(* IEC 61131-3 sources: kkh_knowHow_dgtt/tools/fmse/plc_lib (part 2) *)

(* ---- FB_SafetyCoupling.st ---- *)
(*==================================================================================================================
  FB_SafetyCoupling  -  safety coupling to the neighbour module (e-stop in + zone free)
  ----------------------------------------------------------------------------------------------------------------
  Library   : FMSE device FB library (item 10A)              Version : 1.0.0 (2026-11-15)
  Rule      : tools/fmse/examples/item10a_examples.json  _rules.fb_library (= 2 x FB_Safe2Ch)
  Codegen   : item 8 pattern COUPLING -> st_codegen.py calls this FB (x<Signal> / q<Signal>)
  Purpose   : Item 8 COUPLING: one FB_Safe2Ch for the e-stop chain coming in, one for the zone-free signal of
              the neighbour. The outputs EstopOut / EnableOut are F-outputs written only by the F-program.
  Interface :
    dir  name                type          default   meaning
    IN   xEstopIn            BOOL          -         e-stop in channel 1 F-copy
    IN   xEstopIn2           BOOL          -         e-stop in channel 2 F-copy
    IN   xZoneFree           BOOL          -         zone free channel 1 F-copy
    IN   xZoneFree2          BOOL          -         zone free channel 2 F-copy
    IN   xReset              BOOL          -         fault reset, rising edge
    CFG  tDisc_ms            DINT          500       discrepancy time [ms]
    OUT  xEstopOk            BOOL          -         e-stop chain closed and reset
    OUT  xZoneOk             BOOL          -         neighbour zone free and reset
    OUT  xResetReq           BOOL          -         one of the two waits for a reset
    OUT  xDiscErr            BOOL          -         discrepancy in one of the two
    OUT  iAlarm              INT           -         local alarm code (0 = none)
  Alarms    : iAlarm = local code a ; Admin.AlarmNo = M*1000 + 10*i + a (decision D2), class per module (D3)
    1  e-stop coupling discrepancy
    2  zone-free coupling discrepancy
  Timing    : Times are counted in calls: n * GC_CYCLE_MS >= t_ms (GC_CYCLE_MS = 100 ms = test bench, TYPES.st).
              In the 10 ms main task set GC_CYCLE_MS := 10 (same behaviour, 10 ms resolution) or replace a counter
              by a TON: ton(IN := <condition>, PT := T#2s); IF ton.Q THEN ... (one call later than the counter).
  Siemens   : SCL (TIA Portal): the same statements; local names are written with '#' (#xRst), the VAR section is
              VAR (STAT) of an FB with an instance DB, R_TRIG / TON are multi-instances, enumerations become INT
              constants (E_DriveState.FAULT -> 9), MIN / LIMIT exist, '16#0080' is written W#16#80 for a WORD.
  NOTICE    : ALL VALUES ARE EXAMPLES. Real PLC code is written, reviewed, tested and signed off by qualified
              people. Safety functions only in the F-program; this FB only reads F-copies and writes no F-signal.
==================================================================================================================*)
FUNCTION_BLOCK FB_SafetyCoupling
VAR_INPUT  (* signals *)
  xEstopIn : BOOL;                          (* e-stop in channel 1 F-copy *)
  xEstopIn2 : BOOL;                         (* e-stop in channel 2 F-copy *)
  xZoneFree : BOOL;                         (* zone free channel 1 F-copy *)
  xZoneFree2 : BOOL;                        (* zone free channel 2 F-copy *)
  xReset : BOOL;                            (* fault reset, rising edge *)
END_VAR
VAR_INPUT  (* configuration (set once, defaults = example values) *)
  tDisc_ms : DINT := 500;                   (* discrepancy time [ms] *)
END_VAR
VAR_OUTPUT  (* outputs *)
  xEstopOk : BOOL;                          (* e-stop chain closed and reset *)
  xZoneOk : BOOL;                           (* neighbour zone free and reset *)
  xResetReq : BOOL;                         (* one of the two waits for a reset *)
  xDiscErr : BOOL;                          (* discrepancy in one of the two *)
  iAlarm : INT;                             (* local alarm code (0 = none) *)
END_VAR
VAR  (* internal *)
  fbEstop : FB_Safe2Ch;                     (* e-stop in *)
  fbZone : FB_Safe2Ch;                      (* zone free *)
END_VAR
fbEstop(xCh1 := xEstopIn, xCh2 := xEstopIn2, xReset := xReset, tDisc_ms := tDisc_ms);
fbZone(xCh1 := xZoneFree, xCh2 := xZoneFree2, xReset := xReset, tDisc_ms := tDisc_ms);
xEstopOk := fbEstop.xOk;
xZoneOk := fbZone.xOk;
xResetReq := fbEstop.xResetReq OR fbZone.xResetReq;
xDiscErr := fbEstop.xDiscErr OR fbZone.xDiscErr;
IF fbEstop.xDiscErr THEN
  iAlarm := 1;                                (* e-stop coupling discrepancy *)
ELSIF fbZone.xDiscErr THEN
  iAlarm := 2;                                (* zone-free coupling discrepancy *)
ELSE
  iAlarm := 0;
END_IF
END_FUNCTION_BLOCK

(* ---- FB_SafeValve.st ---- *)
(*==================================================================================================================
  FB_SafeValve  -  redundant safety valve pair with position feedback
  ----------------------------------------------------------------------------------------------------------------
  Library   : FMSE device FB library (item 10A)              Version : 1.0.0 (2026-11-15)
  Rule      : tools/fmse/examples/item10a_examples.json  _rules.fb_library (= 2 x FB_Edm, bInverted FALSE)
  Codegen   : item 8 pattern SAFE_VALVE -> st_codegen.py calls this FB (x<Signal> / q<Signal>)
  Purpose   : Item 8 SAFE_VALVE: two valves (F-outputs ValveA / ValveB written only by the F-program), each
              with a position switch TRUE = open; FB_Edm with bInverted FALSE checks that each follows.
  Interface :
    dir  name                type          default   meaning
    IN   xCmdA               BOOL          -         F-copy of the F-output ValveA
    IN   xCmdB               BOOL          -         F-copy of the F-output ValveB
    IN   xFbA                BOOL          -         valve A open (DI)
    IN   xFbB                BOOL          -         valve B open (DI)
    IN   xReset              BOOL          -         fault reset, rising edge
    CFG  tEdm_ms             DINT          300       feedback time [ms]
    OUT  xOnA                BOOL          -         valve A open and feedback ok
    OUT  xOnB                BOOL          -         valve B open and feedback ok
    OUT  xError              BOOL          -         error latched (see alarms)
    OUT  iAlarm              INT           -         local alarm code (0 = none)
  Alarms    : iAlarm = local code a ; Admin.AlarmNo = M*1000 + 10*i + a (decision D2), class per module (D3)
    1  valve A feedback does not follow
    2  valve B feedback does not follow
  Timing    : Times are counted in calls: n * GC_CYCLE_MS >= t_ms (GC_CYCLE_MS = 100 ms = test bench, TYPES.st).
              In the 10 ms main task set GC_CYCLE_MS := 10 (same behaviour, 10 ms resolution) or replace a counter
              by a TON: ton(IN := <condition>, PT := T#2s); IF ton.Q THEN ... (one call later than the counter).
  Siemens   : SCL (TIA Portal): the same statements; local names are written with '#' (#xRst), the VAR section is
              VAR (STAT) of an FB with an instance DB, R_TRIG / TON are multi-instances, enumerations become INT
              constants (E_DriveState.FAULT -> 9), MIN / LIMIT exist, '16#0080' is written W#16#80 for a WORD.
  NOTICE    : ALL VALUES ARE EXAMPLES. Real PLC code is written, reviewed, tested and signed off by qualified
              people. Safety functions only in the F-program; this FB only reads F-copies and writes no F-signal.
==================================================================================================================*)
FUNCTION_BLOCK FB_SafeValve
VAR_INPUT  (* signals *)
  xCmdA : BOOL;                             (* F-copy of the F-output ValveA *)
  xCmdB : BOOL;                             (* F-copy of the F-output ValveB *)
  xFbA : BOOL;                              (* valve A open (DI) *)
  xFbB : BOOL;                              (* valve B open (DI) *)
  xReset : BOOL;                            (* fault reset, rising edge *)
END_VAR
VAR_INPUT  (* configuration (set once, defaults = example values) *)
  tEdm_ms : DINT := 300;                    (* feedback time [ms] *)
END_VAR
VAR_OUTPUT  (* outputs *)
  xOnA : BOOL;                              (* valve A open and feedback ok *)
  xOnB : BOOL;                              (* valve B open and feedback ok *)
  xError : BOOL;                            (* error latched (see alarms) *)
  iAlarm : INT;                             (* local alarm code (0 = none) *)
END_VAR
VAR  (* internal *)
  fbA : FB_Edm;                             (* EDM valve A *)
  fbB : FB_Edm;                             (* EDM valve B *)
END_VAR
fbA(xCmd := xCmdA, xFb := xFbA, xReset := xReset, tEdm_ms := tEdm_ms, bInverted := FALSE);
fbB(xCmd := xCmdB, xFb := xFbB, xReset := xReset, tEdm_ms := tEdm_ms, bInverted := FALSE);
xOnA := fbA.xOn;
xOnB := fbB.xOn;
xError := fbA.xError OR fbB.xError;
IF fbA.xError THEN
  iAlarm := 1;                                (* valve A feedback *)
ELSIF fbB.xError THEN
  iAlarm := 2;                                (* valve B feedback *)
ELSE
  iAlarm := 0;
END_IF
END_FUNCTION_BLOCK

(* ---- FB_Scanner.st ---- *)
(*==================================================================================================================
  FB_Scanner  -  safety laser scanner: field-set switching and OSSD mirror
  ----------------------------------------------------------------------------------------------------------------
  Library   : FMSE device FB library (item 10A)              Version : 1.0.0 (2026-11-15)
  Rule      : tools/fmse/examples/item10a_examples.json  _rules.FB_Scanner
  Codegen   : item 8 pattern SCANNER -> st_codegen.py calls this FB (x<Signal> / q<Signal>)
  Purpose   : The standard program selects the field set (the scanner checks the combination); the OSSD pair
              and the warning field are mirrored for diagnosis and HMI.
  Interface :
    dir  name                type          default   meaning
    IN   xOssd1              BOOL          -         OSSD 1 F-copy (TRUE = free)
    IN   xOssd2              BOOL          -         OSSD 2 F-copy (TRUE = free)
    IN   xWarn               BOOL          -         warning field interrupted (DI)
    IN   iField              INT           1         field set 1 = A, 2 = B
    OUT  qFieldA             BOOL          -         field set A select (DO)
    OUT  qFieldB             BOOL          -         field set B select (DO)
    OUT  xFree               BOOL          -         protective field free
    OUT  xWarnOut            BOOL          -         warning field interrupted
    OUT  iAlarm              INT           -         local alarm code (0 = none)
  Alarms    : iAlarm = local code a ; Admin.AlarmNo = M*1000 + 10*i + a (decision D2), class per module (D3)
    2  invalid field set
  Timing    : Times are counted in calls: n * GC_CYCLE_MS >= t_ms (GC_CYCLE_MS = 100 ms = test bench, TYPES.st).
              In the 10 ms main task set GC_CYCLE_MS := 10 (same behaviour, 10 ms resolution) or replace a counter
              by a TON: ton(IN := <condition>, PT := T#2s); IF ton.Q THEN ... (one call later than the counter).
  Siemens   : SCL (TIA Portal): the same statements; local names are written with '#' (#xRst), the VAR section is
              VAR (STAT) of an FB with an instance DB, R_TRIG / TON are multi-instances, enumerations become INT
              constants (E_DriveState.FAULT -> 9), MIN / LIMIT exist, '16#0080' is written W#16#80 for a WORD.
  NOTICE    : ALL VALUES ARE EXAMPLES. Real PLC code is written, reviewed, tested and signed off by qualified
              people. Safety functions only in the F-program; this FB only reads F-copies and writes no F-signal.
==================================================================================================================*)
FUNCTION_BLOCK FB_Scanner
VAR_INPUT  (* signals *)
  xOssd1 : BOOL;                            (* OSSD 1 F-copy (TRUE = free) *)
  xOssd2 : BOOL;                            (* OSSD 2 F-copy (TRUE = free) *)
  xWarn : BOOL;                             (* warning field interrupted (DI) *)
  iField : INT := 1;                        (* field set 1 = A, 2 = B *)
END_VAR
VAR_OUTPUT  (* outputs *)
  qFieldA : BOOL;                           (* field set A select (DO) *)
  qFieldB : BOOL;                           (* field set B select (DO) *)
  xFree : BOOL;                             (* protective field free *)
  xWarnOut : BOOL;                          (* warning field interrupted *)
  iAlarm : INT;                             (* local alarm code (0 = none) *)
END_VAR
qFieldA := iField = 1;
qFieldB := iField = 2;
xFree := xOssd1 AND xOssd2;
xWarnOut := xWarn;
IF iField = 1 OR iField = 2 THEN
  iAlarm := 0;
ELSE
  iAlarm := 2;                                (* invalid field set *)
END_IF
END_FUNCTION_BLOCK

(* ---- FB_Sensor.st ---- *)
(*==================================================================================================================
  FB_Sensor  -  digital sensor with on / off debounce
  ----------------------------------------------------------------------------------------------------------------
  Library   : FMSE device FB library (item 10A)              Version : 1.0.0 (2026-11-15)
  Rule      : tools/fmse/examples/item10a_examples.json  _rules.FB_Sensor
  Codegen   : item 8 pattern SENSOR -> st_codegen.py calls this FB (x<Signal> / q<Signal>)
  Purpose   : Debounce of a digital sensor: the value follows the input only after it differs for tOn_ms (0 -> 1)
              or tOff_ms (1 -> 0); a shorter bounce is ignored. tOn_ms = tOff_ms = 0: one call delay is not added.
  Interface :
    dir  name                type          default   meaning
    IN   xOn                 BOOL          -         sensor input (DI)
    CFG  tOn_ms              DINT          0         debounce time 0 -> 1 [ms]
    CFG  tOff_ms             DINT          0         debounce time 1 -> 0 [ms]
    OUT  xValue              BOOL          -         debounced value
  Alarms    : iAlarm = local code a ; Admin.AlarmNo = M*1000 + 10*i + a (decision D2), class per module (D3)
    none
  Timing    : Times are counted in calls: n * GC_CYCLE_MS >= t_ms (GC_CYCLE_MS = 100 ms = test bench, TYPES.st).
              In the 10 ms main task set GC_CYCLE_MS := 10 (same behaviour, 10 ms resolution) or replace a counter
              by a TON: ton(IN := <condition>, PT := T#2s); IF ton.Q THEN ... (one call later than the counter).
  Siemens   : SCL (TIA Portal): the same statements; local names are written with '#' (#xRst), the VAR section is
              VAR (STAT) of an FB with an instance DB, R_TRIG / TON are multi-instances, enumerations become INT
              constants (E_DriveState.FAULT -> 9), MIN / LIMIT exist, '16#0080' is written W#16#80 for a WORD.
  NOTICE    : ALL VALUES ARE EXAMPLES. Real PLC code is written, reviewed, tested and signed off by qualified
              people. Safety functions only in the F-program; this FB only reads F-copies and writes no F-signal.
==================================================================================================================*)
FUNCTION_BLOCK FB_Sensor
VAR_INPUT  (* signals *)
  xOn : BOOL;                               (* sensor input (DI) *)
END_VAR
VAR_INPUT  (* configuration (set once, defaults = example values) *)
  tOn_ms : DINT := 0;                       (* debounce time 0 -> 1 [ms] *)
  tOff_ms : DINT := 0;                      (* debounce time 1 -> 0 [ms] *)
END_VAR
VAR_OUTPUT  (* outputs *)
  xValue : BOOL;                            (* debounced value *)
END_VAR
VAR  (* internal *)
  nCnt : DINT;                              (* calls with input <> value *)
  tLim : DINT;                              (* active debounce time *)
END_VAR
IF xOn <> xValue THEN
  nCnt := MIN(nCnt + 1, GC_N_MAX);
  IF xOn THEN
    tLim := tOn_ms;
  ELSE
    tLim := tOff_ms;
  END_IF
  IF nCnt * GC_CYCLE_MS >= tLim THEN
    xValue := xOn;
    nCnt := 0;
  END_IF
ELSE
  nCnt := 0;
END_IF
END_FUNCTION_BLOCK

(* ---- FB_SignalTower.st ---- *)
(*==================================================================================================================
  FB_SignalTower  -  signal tower (stack light) and horn per PackML state and alarm class
  ----------------------------------------------------------------------------------------------------------------
  Library   : FMSE device FB library (item 10A)              Version : 1.0.0 (2026-11-15)
  Rule      : tools/fmse/examples/item10a_examples.json  _rules.FB_SignalTower
  Codegen   : item 8 pattern SIGNAL_TOWER -> st_codegen.py calls this FB (x<Signal> / q<Signal>)
  Purpose   : Colours per IEC 60204-1 10.3 / IEC 60073: red = class A alarm or Aborting/Aborted, yellow = class
              B/C or Stopped/Suspended/Held, green = running states, flashing green = Idle/Complete (ready).
              Horn on a new class A/B alarm until acknowledged or no alarm.
  Interface :
    dir  name                type          default   meaning
    IN   iState              INT           2         PackML state number (2 = Stopped)
    IN   iAlarmClass         INT           -         0 none, 1 A, 2 B, 3 C (FB_AlarmMgr)
    IN   xHornAck            BOOL          -         horn acknowledge, rising edge
    OUT  qRed                BOOL          -         red lamp (DO)
    OUT  qYellow             BOOL          -         yellow lamp (DO)
    OUT  qGreen              BOOL          -         green lamp (DO)
    OUT  qBuzzer             BOOL          -         horn (DO)
  Alarms    : iAlarm = local code a ; Admin.AlarmNo = M*1000 + 10*i + a (decision D2), class per module (D3)
    none
  Timing    : Times are counted in calls: n * GC_CYCLE_MS >= t_ms (GC_CYCLE_MS = 100 ms = test bench, TYPES.st).
              In the 10 ms main task set GC_CYCLE_MS := 10 (same behaviour, 10 ms resolution) or replace a counter
              by a TON: ton(IN := <condition>, PT := T#2s); IF ton.Q THEN ... (one call later than the counter).
  Siemens   : SCL (TIA Portal): the same statements; local names are written with '#' (#xRst), the VAR section is
              VAR (STAT) of an FB with an instance DB, R_TRIG / TON are multi-instances, enumerations become INT
              constants (E_DriveState.FAULT -> 9), MIN / LIMIT exist, '16#0080' is written W#16#80 for a WORD.
  NOTICE    : ALL VALUES ARE EXAMPLES. Real PLC code is written, reviewed, tested and signed off by qualified
              people. Safety functions only in the F-program; this FB only reads F-copies and writes no F-signal.
==================================================================================================================*)
FUNCTION_BLOCK FB_SignalTower
VAR_INPUT  (* signals *)
  iState : INT := 2;                        (* PackML state number (2 = Stopped) *)
  iAlarmClass : INT;                        (* 0 none, 1 A, 2 B, 3 C (FB_AlarmMgr) *)
  xHornAck : BOOL;                          (* horn acknowledge, rising edge *)
END_VAR
VAR_OUTPUT  (* outputs *)
  qRed : BOOL;                              (* red lamp (DO) *)
  qYellow : BOOL;                           (* yellow lamp (DO) *)
  qGreen : BOOL;                            (* green lamp (DO) *)
  qBuzzer : BOOL;                           (* horn (DO) *)
END_VAR
VAR  (* internal *)
  nBlink : DINT;                            (* blink counter 0 .. 2*nHalf-1 *)
  nHalf : DINT;                             (* calls per half period *)
  xBlink : BOOL;                            (* 1 Hz blink, TRUE in the first half *)
  rtAck : R_TRIG;                           (* edge of xHornAck *)
  iPrevClass : INT;                         (* alarm class of the last call *)
  xHorn : BOOL;                             (* horn latch *)
END_VAR
nHalf := GC_BLINK_HALF_MS / GC_CYCLE_MS;     (* 5 calls at 100 ms = 1 Hz *)
xBlink := nBlink < nHalf;
nBlink := (nBlink + 1) MOD (2 * nHalf);
rtAck(CLK := xHornAck);
qRed := (iAlarmClass = E_AlarmClass.A) OR (iState = E_PackMLState.ABORTING) OR (iState = E_PackMLState.ABORTED);
qYellow := (iAlarmClass = E_AlarmClass.B) OR (iAlarmClass = E_AlarmClass.C) OR (iState = E_PackMLState.STOPPED)
           OR (iState = E_PackMLState.SUSPENDED) OR (iState = E_PackMLState.HELD);
CASE iState OF
  E_PackMLState.STARTING, E_PackMLState.EXECUTE, E_PackMLState.UNHOLDING, E_PackMLState.UNSUSPENDING,
  E_PackMLState.COMPLETING:
    qGreen := TRUE;
  E_PackMLState.IDLE, E_PackMLState.COMPLETE:
    qGreen := xBlink;                         (* flashing green = ready, waiting *)
ELSE
  qGreen := FALSE;
END_CASE
IF (iAlarmClass = E_AlarmClass.A OR iAlarmClass = E_AlarmClass.B) AND iAlarmClass <> iPrevClass THEN
  xHorn := TRUE;
END_IF
IF rtAck.Q OR iAlarmClass = E_AlarmClass.NONE THEN
  xHorn := FALSE;
END_IF
iPrevClass := iAlarmClass;
qBuzzer := xHorn;
END_FUNCTION_BLOCK

(* ---- FB_TwoHand.st ---- *)
(*==================================================================================================================
  FB_TwoHand  -  diagnostic mirror of a two-hand control (type IIIC)
  ----------------------------------------------------------------------------------------------------------------
  Library   : FMSE device FB library (item 10A)              Version : 1.0.0 (2026-11-15)
  Rule      : tools/fmse/examples/item10a_examples.json  _rules.FB_TwoHand
  Codegen   : item 8 pattern TWOHAND -> st_codegen.py calls this FB (x<Signal> / q<Signal>)
  Purpose   : Two 2-channel buttons, simultaneity 0.5 s (the F-program does the safety function). Pressing the
              second hand later than tSync_ms blocks until both are released. Strict '>': the 5th call (500 ms)
              is still simultaneous.
  Interface :
    dir  name                type          default   meaning
    IN   xLeft               BOOL          -         left button NO (DI)
    IN   xLeft2              BOOL          -         left button NC (DI)
    IN   xRight              BOOL          -         right button NO (DI)
    IN   xRight2             BOOL          -         right button NC (DI)
    CFG  tSync_ms            DINT          500       simultaneity time [ms]
    OUT  xActuated           BOOL          -         both hands, simultaneous
    OUT  xError              BOOL          -         error latched (see alarms)
    OUT  iAlarm              INT           -         local alarm code (0 = none)
  Alarms    : iAlarm = local code a ; Admin.AlarmNo = M*1000 + 10*i + a (decision D2), class per module (D3)
    1  not simultaneous - release both
  Timing    : Times are counted in calls: n * GC_CYCLE_MS >= t_ms (GC_CYCLE_MS = 100 ms = test bench, TYPES.st).
              In the 10 ms main task set GC_CYCLE_MS := 10 (same behaviour, 10 ms resolution) or replace a counter
              by a TON: ton(IN := <condition>, PT := T#2s); IF ton.Q THEN ... (one call later than the counter).
  Siemens   : SCL (TIA Portal): the same statements; local names are written with '#' (#xRst), the VAR section is
              VAR (STAT) of an FB with an instance DB, R_TRIG / TON are multi-instances, enumerations become INT
              constants (E_DriveState.FAULT -> 9), MIN / LIMIT exist, '16#0080' is written W#16#80 for a WORD.
  NOTICE    : ALL VALUES ARE EXAMPLES. Real PLC code is written, reviewed, tested and signed off by qualified
              people. Safety functions only in the F-program; this FB only reads F-copies and writes no F-signal.
==================================================================================================================*)
FUNCTION_BLOCK FB_TwoHand
VAR_INPUT  (* signals *)
  xLeft : BOOL;                             (* left button NO (DI) *)
  xLeft2 : BOOL;                            (* left button NC (DI) *)
  xRight : BOOL;                            (* right button NO (DI) *)
  xRight2 : BOOL;                           (* right button NC (DI) *)
END_VAR
VAR_INPUT  (* configuration (set once, defaults = example values) *)
  tSync_ms : DINT := 500;                   (* simultaneity time [ms] *)
END_VAR
VAR_OUTPUT  (* outputs *)
  xActuated : BOOL;                         (* both hands, simultaneous *)
  xError : BOOL;                            (* error latched (see alarms) *)
  iAlarm : INT;                             (* local alarm code (0 = none) *)
END_VAR
VAR  (* internal *)
  xL : BOOL;                                (* left actuated *)
  xR : BOOL;                                (* right actuated *)
  n : DINT;                                 (* calls with one hand only *)
  xBlocked : BOOL;                          (* release both first *)
END_VAR
xL := xLeft AND xLeft2;
xR := xRight AND xRight2;
IF NOT xL AND NOT xR THEN
  xBlocked := FALSE;
  n := 0;
  xError := FALSE;
  iAlarm := 0;
  xActuated := FALSE;
ELSIF xL <> xR THEN
  n := MIN(n + 1, GC_N_MAX);
  IF (n * GC_CYCLE_MS > tSync_ms) AND NOT xActuated THEN
    xBlocked := TRUE;
    xError := TRUE;
    iAlarm := 1;                              (* not simultaneous *)
  END_IF
  xActuated := FALSE;
ELSE
  xActuated := NOT xBlocked;
END_IF
END_FUNCTION_BLOCK

(* ---- FB_Ups.st ---- *)
(*==================================================================================================================
  FB_Ups  -  24 V DC UPS monitoring with shutdown request
  ----------------------------------------------------------------------------------------------------------------
  Library   : FMSE device FB library (item 10A)              Version : 1.0.0 (2026-11-15)
  Rule      : tools/fmse/examples/item10a_examples.json  _rules.FB_Ups
  Codegen   : item 8 pattern UPS_DC -> st_codegen.py calls this FB (x<Signal> / q<Signal>)
  Purpose   : UPS signals: fault, on battery; after tBuffer_ms on battery the PLC / PC shut down in order.
  Interface :
    dir  name                type          default   meaning
    IN   xUpsOk              BOOL          TRUE      UPS ready / no fault (DI)
    IN   xOnBattery          BOOL          -         mains lost, on battery (DI)
    CFG  tBuffer_ms          DINT          5000      buffer time before shutdown [ms]
    OUT  xShutdownReq        BOOL          -         request an orderly shutdown
    OUT  iAlarm              INT           -         local alarm code (0 = none)
  Alarms    : iAlarm = local code a ; Admin.AlarmNo = M*1000 + 10*i + a (decision D2), class per module (D3)
    1  UPS fault
    2  on battery
  Timing    : Times are counted in calls: n * GC_CYCLE_MS >= t_ms (GC_CYCLE_MS = 100 ms = test bench, TYPES.st).
              In the 10 ms main task set GC_CYCLE_MS := 10 (same behaviour, 10 ms resolution) or replace a counter
              by a TON: ton(IN := <condition>, PT := T#2s); IF ton.Q THEN ... (one call later than the counter).
  Siemens   : SCL (TIA Portal): the same statements; local names are written with '#' (#xRst), the VAR section is
              VAR (STAT) of an FB with an instance DB, R_TRIG / TON are multi-instances, enumerations become INT
              constants (E_DriveState.FAULT -> 9), MIN / LIMIT exist, '16#0080' is written W#16#80 for a WORD.
  NOTICE    : ALL VALUES ARE EXAMPLES. Real PLC code is written, reviewed, tested and signed off by qualified
              people. Safety functions only in the F-program; this FB only reads F-copies and writes no F-signal.
==================================================================================================================*)
FUNCTION_BLOCK FB_Ups
VAR_INPUT  (* signals *)
  xUpsOk : BOOL := TRUE;                    (* UPS ready / no fault (DI) *)
  xOnBattery : BOOL;                        (* mains lost, on battery (DI) *)
END_VAR
VAR_INPUT  (* configuration (set once, defaults = example values) *)
  tBuffer_ms : DINT := 5000;                (* buffer time before shutdown [ms] *)
END_VAR
VAR_OUTPUT  (* outputs *)
  xShutdownReq : BOOL;                      (* request an orderly shutdown *)
  iAlarm : INT;                             (* local alarm code (0 = none) *)
END_VAR
VAR  (* internal *)
  n : DINT;                                 (* calls on battery *)
END_VAR
IF xOnBattery THEN
  n := MIN(n + 1, GC_N_MAX);
ELSE
  n := 0;
END_IF
xShutdownReq := n * GC_CYCLE_MS >= tBuffer_ms;
IF NOT xUpsOk THEN
  iAlarm := 1;                                (* UPS fault *)
ELSIF xOnBattery THEN
  iAlarm := 2;                                (* on battery *)
ELSE
  iAlarm := 0;
END_IF
END_FUNCTION_BLOCK

(* ---- FB_Valve1.st ---- *)
(*==================================================================================================================
  FB_Valve1  -  single-solenoid valve (spring return) with end-position monitoring
  ----------------------------------------------------------------------------------------------------------------
  Library   : FMSE device FB library (item 10A)              Version : 1.0.0 (2026-11-15)
  Rule      : tools/fmse/examples/item10a_examples.json  _rules.FB_Valve
  Codegen   : item 8 pattern VALVE_SINGLE -> st_codegen.py calls this FB (x<Signal> / q<Signal>)
  Purpose   : Pneumatic cylinder with a 5/2 single-solenoid valve: qSol TRUE -> position B, FALSE (or xEnable
              FALSE) -> the spring returns it to A. Supervises the movement time, the loss of the end position and
              both end switches; a reset retries the movement.
  Interface :
    dir  name                type          default   meaning
    IN   xPosA               BOOL          TRUE      end switch A (DI); default: starts at A
    IN   xPosB               BOOL          -         end switch B (DI)
    IN   xCmdB               BOOL          -         TRUE = go to / stay at B, FALSE = A
    IN   xEnable             BOOL          TRUE      FALSE = outputs off
    IN   xReset              BOOL          -         fault reset, rising edge
    CFG  tMove_ms            DINT          2000      max. time to reach the end position [ms]
    CFG  tLost_ms            DINT          300       end position lost without command [ms]
    CFG  tBoth_ms            DINT          200       both end switches on [ms]
    OUT  qSol                BOOL          -         solenoid (DO): TRUE = B
    OUT  xAtA                BOOL          -         at end position A
    OUT  xAtB                BOOL          -         at end position B
    OUT  xBusy               BOOL          -         moving (supervised)
    OUT  xError              BOOL          -         error latched (see alarms)
    OUT  iAlarm              INT           -         local alarm code (0 = none)
  Alarms    : iAlarm = local code a ; Admin.AlarmNo = M*1000 + 10*i + a (decision D2), class per module (D3)
    1  end position not reached
    2  left the end position without command
    3  both end switches on
  Timing    : Times are counted in calls: n * GC_CYCLE_MS >= t_ms (GC_CYCLE_MS = 100 ms = test bench, TYPES.st).
              In the 10 ms main task set GC_CYCLE_MS := 10 (same behaviour, 10 ms resolution) or replace a counter
              by a TON: ton(IN := <condition>, PT := T#2s); IF ton.Q THEN ... (one call later than the counter).
  Siemens   : SCL (TIA Portal): the same statements; local names are written with '#' (#xRst), the VAR section is
              VAR (STAT) of an FB with an instance DB, R_TRIG / TON are multi-instances, enumerations become INT
              constants (E_DriveState.FAULT -> 9), MIN / LIMIT exist, '16#0080' is written W#16#80 for a WORD.
  NOTICE    : ALL VALUES ARE EXAMPLES. Real PLC code is written, reviewed, tested and signed off by qualified
              people. Safety functions only in the F-program; this FB only reads F-copies and writes no F-signal.
==================================================================================================================*)
FUNCTION_BLOCK FB_Valve1
VAR_INPUT  (* signals *)
  xPosA : BOOL := TRUE;                     (* end switch A (DI); default: starts at A *)
  xPosB : BOOL;                             (* end switch B (DI) *)
  xCmdB : BOOL;                             (* TRUE = go to / stay at B, FALSE = A *)
  xEnable : BOOL := TRUE;                   (* FALSE = outputs off *)
  xReset : BOOL;                            (* fault reset, rising edge *)
END_VAR
VAR_INPUT  (* configuration (set once, defaults = example values) *)
  tMove_ms : DINT := 2000;                  (* max. time to reach the end position [ms] *)
  tLost_ms : DINT := 300;                   (* end position lost without command [ms] *)
  tBoth_ms : DINT := 200;                   (* both end switches on [ms] *)
END_VAR
VAR_OUTPUT  (* outputs *)
  qSol : BOOL;                              (* solenoid (DO): TRUE = B *)
  xAtA : BOOL;                              (* at end position A *)
  xAtB : BOOL;                              (* at end position B *)
  xBusy : BOOL;                             (* moving (supervised) *)
  xError : BOOL;                            (* error latched (see alarms) *)
  iAlarm : INT;                             (* local alarm code (0 = none) *)
END_VAR
VAR  (* internal *)
  rtReset : R_TRIG;                         (* edge of xReset *)
  xRst : BOOL;                              (* reset pulse *)
  xA : BOOL;                                (* at A (decoded) *)
  xB : BOOL;                                (* at B (decoded) *)
  xReached : BOOL;                          (* commanded end position reached *)
  xMoving : BOOL;                           (* movement supervised *)
  xPrevCmd : BOOL;                          (* command of the last call *)
  xFirst : BOOL := TRUE;                    (* first call *)
  nMove : DINT;                             (* calls while moving and enabled *)
  nLost : DINT;                             (* calls out of position *)
  nBoth : DINT;                             (* calls with both switches on *)
END_VAR
(* step 0: edge of the reset and position decode *)
rtReset(CLK := xReset);
xRst := rtReset.Q;
xA := xPosA AND NOT xPosB;
xB := xPosB AND NOT xPosA;
IF xCmdB THEN
  xReached := xB;
ELSE
  xReached := xA;
END_IF
(* (1) reset of an error = retry: supervise the movement again if the end position is not reached *)
IF xError AND xRst AND NOT (xPosA AND xPosB) THEN
  xError := FALSE;
  iAlarm := 0;
  xMoving := NOT xReached;
  nMove := 0;
  nLost := 0;
END_IF
(* (2) new command or first call: start the movement supervision *)
IF xFirst OR (xCmdB <> xPrevCmd) THEN
  xMoving := TRUE;
  nMove := 0;
END_IF
(* (3) both end switches on at the same time *)
IF xPosA AND xPosB THEN
  nBoth := MIN(nBoth + 1, GC_N_MAX);
ELSE
  nBoth := 0;
END_IF
(* (4) supervision - an error latches until a reset *)
IF NOT xError THEN
  IF nBoth * GC_CYCLE_MS >= tBoth_ms THEN
    xError := TRUE;
    iAlarm := 3;                              (* both end switches on *)
    xMoving := FALSE;
  ELSIF xMoving THEN
    nLost := 0;
    IF xEnable THEN                           (* the movement timer pauses while disabled *)
      nMove := MIN(nMove + 1, GC_N_MAX);
      IF xReached THEN
        xMoving := FALSE;
      ELSIF nMove * GC_CYCLE_MS >= tMove_ms THEN
        xError := TRUE;
        iAlarm := 1;                          (* end position not reached *)
        xMoving := FALSE;
      END_IF
    END_IF
  ELSIF xEnable THEN
    IF NOT xReached THEN
      nLost := MIN(nLost + 1, GC_N_MAX);
    ELSE
      nLost := 0;
    END_IF
    IF nLost * GC_CYCLE_MS >= tLost_ms THEN
      xError := TRUE;
      iAlarm := 2;                            (* left the end position without command *)
    END_IF
  ELSE
    nLost := 0;
  END_IF
END_IF
(* (5) outputs - an error does NOT switch the solenoid(s): the module reacts by alarm class (D3) *)
qSol := xCmdB AND xEnable;
xAtA := xA;
xAtB := xB;
xBusy := xMoving AND NOT xError;
xPrevCmd := xCmdB;
xFirst := FALSE;
END_FUNCTION_BLOCK

(* ---- FB_Valve2.st ---- *)
(*==================================================================================================================
  FB_Valve2  -  double-solenoid (bistable) valve with end-position monitoring
  ----------------------------------------------------------------------------------------------------------------
  Library   : FMSE device FB library (item 10A)              Version : 1.0.0 (2026-11-15)
  Rule      : tools/fmse/examples/item10a_examples.json  _rules.FB_Valve
  Codegen   : item 8 pattern VALVE_DOUBLE -> st_codegen.py calls this FB (x<Signal> / q<Signal>)
  Purpose   : Pneumatic cylinder / rotary actuator with a 5/2 double-solenoid valve: qSolB drives to B, qSolA to A.
              xEnable FALSE switches both solenoids off and the valve HOLDS its position (the movement timer
              pauses). Same supervision and alarms as FB_Valve1.
  Interface :
    dir  name                type          default   meaning
    IN   xPosA               BOOL          TRUE      end switch A (DI); default: starts at A
    IN   xPosB               BOOL          -         end switch B (DI)
    IN   xCmdB               BOOL          -         TRUE = go to / stay at B, FALSE = A
    IN   xEnable             BOOL          TRUE      FALSE = outputs off
    IN   xReset              BOOL          -         fault reset, rising edge
    CFG  tMove_ms            DINT          2000      max. time to reach the end position [ms]
    CFG  tLost_ms            DINT          300       end position lost without command [ms]
    CFG  tBoth_ms            DINT          200       both end switches on [ms]
    OUT  qSolA               BOOL          -         solenoid A (DO)
    OUT  qSolB               BOOL          -         solenoid B (DO)
    OUT  xAtA                BOOL          -         at end position A
    OUT  xAtB                BOOL          -         at end position B
    OUT  xBusy               BOOL          -         moving (supervised)
    OUT  xError              BOOL          -         error latched (see alarms)
    OUT  iAlarm              INT           -         local alarm code (0 = none)
  Alarms    : iAlarm = local code a ; Admin.AlarmNo = M*1000 + 10*i + a (decision D2), class per module (D3)
    1  end position not reached
    2  left the end position without command
    3  both end switches on
  Timing    : Times are counted in calls: n * GC_CYCLE_MS >= t_ms (GC_CYCLE_MS = 100 ms = test bench, TYPES.st).
              In the 10 ms main task set GC_CYCLE_MS := 10 (same behaviour, 10 ms resolution) or replace a counter
              by a TON: ton(IN := <condition>, PT := T#2s); IF ton.Q THEN ... (one call later than the counter).
  Siemens   : SCL (TIA Portal): the same statements; local names are written with '#' (#xRst), the VAR section is
              VAR (STAT) of an FB with an instance DB, R_TRIG / TON are multi-instances, enumerations become INT
              constants (E_DriveState.FAULT -> 9), MIN / LIMIT exist, '16#0080' is written W#16#80 for a WORD.
  NOTICE    : ALL VALUES ARE EXAMPLES. Real PLC code is written, reviewed, tested and signed off by qualified
              people. Safety functions only in the F-program; this FB only reads F-copies and writes no F-signal.
==================================================================================================================*)
FUNCTION_BLOCK FB_Valve2
VAR_INPUT  (* signals *)
  xPosA : BOOL := TRUE;                     (* end switch A (DI); default: starts at A *)
  xPosB : BOOL;                             (* end switch B (DI) *)
  xCmdB : BOOL;                             (* TRUE = go to / stay at B, FALSE = A *)
  xEnable : BOOL := TRUE;                   (* FALSE = outputs off *)
  xReset : BOOL;                            (* fault reset, rising edge *)
END_VAR
VAR_INPUT  (* configuration (set once, defaults = example values) *)
  tMove_ms : DINT := 2000;                  (* max. time to reach the end position [ms] *)
  tLost_ms : DINT := 300;                   (* end position lost without command [ms] *)
  tBoth_ms : DINT := 200;                   (* both end switches on [ms] *)
END_VAR
VAR_OUTPUT  (* outputs *)
  qSolA : BOOL;                             (* solenoid A (DO) *)
  qSolB : BOOL;                             (* solenoid B (DO) *)
  xAtA : BOOL;                              (* at end position A *)
  xAtB : BOOL;                              (* at end position B *)
  xBusy : BOOL;                             (* moving (supervised) *)
  xError : BOOL;                            (* error latched (see alarms) *)
  iAlarm : INT;                             (* local alarm code (0 = none) *)
END_VAR
VAR  (* internal *)
  rtReset : R_TRIG;                         (* edge of xReset *)
  xRst : BOOL;                              (* reset pulse *)
  xA : BOOL;                                (* at A (decoded) *)
  xB : BOOL;                                (* at B (decoded) *)
  xReached : BOOL;                          (* commanded end position reached *)
  xMoving : BOOL;                           (* movement supervised *)
  xPrevCmd : BOOL;                          (* command of the last call *)
  xFirst : BOOL := TRUE;                    (* first call *)
  nMove : DINT;                             (* calls while moving and enabled *)
  nLost : DINT;                             (* calls out of position *)
  nBoth : DINT;                             (* calls with both switches on *)
END_VAR
(* step 0: edge of the reset and position decode *)
rtReset(CLK := xReset);
xRst := rtReset.Q;
xA := xPosA AND NOT xPosB;
xB := xPosB AND NOT xPosA;
IF xCmdB THEN
  xReached := xB;
ELSE
  xReached := xA;
END_IF
(* (1) reset of an error = retry: supervise the movement again if the end position is not reached *)
IF xError AND xRst AND NOT (xPosA AND xPosB) THEN
  xError := FALSE;
  iAlarm := 0;
  xMoving := NOT xReached;
  nMove := 0;
  nLost := 0;
END_IF
(* (2) new command or first call: start the movement supervision *)
IF xFirst OR (xCmdB <> xPrevCmd) THEN
  xMoving := TRUE;
  nMove := 0;
END_IF
(* (3) both end switches on at the same time *)
IF xPosA AND xPosB THEN
  nBoth := MIN(nBoth + 1, GC_N_MAX);
ELSE
  nBoth := 0;
END_IF
(* (4) supervision - an error latches until a reset *)
IF NOT xError THEN
  IF nBoth * GC_CYCLE_MS >= tBoth_ms THEN
    xError := TRUE;
    iAlarm := 3;                              (* both end switches on *)
    xMoving := FALSE;
  ELSIF xMoving THEN
    nLost := 0;
    IF xEnable THEN                           (* the movement timer pauses while disabled *)
      nMove := MIN(nMove + 1, GC_N_MAX);
      IF xReached THEN
        xMoving := FALSE;
      ELSIF nMove * GC_CYCLE_MS >= tMove_ms THEN
        xError := TRUE;
        iAlarm := 1;                          (* end position not reached *)
        xMoving := FALSE;
      END_IF
    END_IF
  ELSIF xEnable THEN
    IF NOT xReached THEN
      nLost := MIN(nLost + 1, GC_N_MAX);
    ELSE
      nLost := 0;
    END_IF
    IF nLost * GC_CYCLE_MS >= tLost_ms THEN
      xError := TRUE;
      iAlarm := 2;                            (* left the end position without command *)
    END_IF
  ELSE
    nLost := 0;
  END_IF
END_IF
(* (5) outputs - an error does NOT switch the solenoid(s): the module reacts by alarm class (D3) *)
qSolB := xCmdB AND xEnable;
qSolA := NOT xCmdB AND xEnable;
xAtA := xA;
xAtB := xB;
xBusy := xMoving AND NOT xError;
xPrevCmd := xCmdB;
xFirst := FALSE;
END_FUNCTION_BLOCK

(* ---- FB_ZoneOut.st ---- *)
(*==================================================================================================================
  FB_ZoneOut  -  safety zone output (released contactors) with EDM
  ----------------------------------------------------------------------------------------------------------------
  Library   : FMSE device FB library (item 10A)              Version : 1.0.0 (2026-11-15)
  Rule      : tools/fmse/examples/item10a_examples.json  _rules.fb_library (= FB_Edm, bInverted TRUE)
  Codegen   : item 8 pattern ZONE_OUT -> st_codegen.py calls this FB (x<Signal> / q<Signal>)
  Purpose   : Wrapper of FB_Edm with bInverted TRUE. The F-output Release is written only by the F-program;
              xCmd is its read-only F-copy.
  Interface :
    dir  name                type          default   meaning
    IN   xCmd                BOOL          -         F-copy of the F-output Release
    IN   xFb                 BOOL          TRUE      NC mirror contacts in series (DI), TRUE = open
    IN   xReset              BOOL          -         fault reset, rising edge
    CFG  tEdm_ms             DINT          300       feedback time [ms]
    OUT  xOn                 BOOL          -         output on and feedback ok
    OUT  xError              BOOL          -         error latched (see alarms)
    OUT  iAlarm              INT           -         local alarm code (0 = none)
  Alarms    : iAlarm = local code a ; Admin.AlarmNo = M*1000 + 10*i + a (decision D2), class per module (D3)
    1  feedback does not follow (welded / not switching)
  Timing    : Times are counted in calls: n * GC_CYCLE_MS >= t_ms (GC_CYCLE_MS = 100 ms = test bench, TYPES.st).
              In the 10 ms main task set GC_CYCLE_MS := 10 (same behaviour, 10 ms resolution) or replace a counter
              by a TON: ton(IN := <condition>, PT := T#2s); IF ton.Q THEN ... (one call later than the counter).
  Siemens   : SCL (TIA Portal): the same statements; local names are written with '#' (#xRst), the VAR section is
              VAR (STAT) of an FB with an instance DB, R_TRIG / TON are multi-instances, enumerations become INT
              constants (E_DriveState.FAULT -> 9), MIN / LIMIT exist, '16#0080' is written W#16#80 for a WORD.
  NOTICE    : ALL VALUES ARE EXAMPLES. Real PLC code is written, reviewed, tested and signed off by qualified
              people. Safety functions only in the F-program; this FB only reads F-copies and writes no F-signal.
==================================================================================================================*)
FUNCTION_BLOCK FB_ZoneOut
VAR_INPUT  (* signals *)
  xCmd : BOOL;                              (* F-copy of the F-output Release *)
  xFb : BOOL := TRUE;                       (* NC mirror contacts in series (DI), TRUE = open *)
  xReset : BOOL;                            (* fault reset, rising edge *)
END_VAR
VAR_INPUT  (* configuration (set once, defaults = example values) *)
  tEdm_ms : DINT := 300;                    (* feedback time [ms] *)
END_VAR
VAR_OUTPUT  (* outputs *)
  xOn : BOOL;                               (* output on and feedback ok *)
  xError : BOOL;                            (* error latched (see alarms) *)
  iAlarm : INT;                             (* local alarm code (0 = none) *)
END_VAR
VAR  (* internal *)
  fbEdm : FB_Edm;                           (* EDM *)
END_VAR
fbEdm(xCmd := xCmd, xFb := xFb, xReset := xReset, tEdm_ms := tEdm_ms, bInverted := TRUE);
xOn := fbEdm.xOn;
xError := fbEdm.xError;
iAlarm := fbEdm.iAlarm;
END_FUNCTION_BLOCK
